Fanuc KAREL source: KA00098.KL

PROGRAM KA00098
%NOLOCKGROUP
VAR
  SRC: VECTOR
  DST: REAL
BEGIN
  SRC.X = 1.0
  DST = SRC
END KA00098
